(* IEC 61131-3 sources: plcassist-cli/packages/volt-lsp-iec/test-corpus/lenze-mid/Device/Plc Logic/Application/Library Manager/CAA MemBlockMan, 91 files *)

(* ---- RSHANDLING.gvl ---- *)
VAR_GLOBAL
	G_XCHGCLASS : XChgClass;
	G_FLATCLASS : FlatClass;
	G_MSGCLASS : MsgClass;
	G_REFCLASS : MsgClass;
	G_POOLCLASS : PoolClass;
	G_BLKCLASS : BlkClass;
	G_RLSTCLASS : RLstClass;
END_VAR

(* ---- VERSIONCONSTANTS.gvl ---- *)
VAR_GLOBAL
	GC_BYVERSION : BYTE := 1;
	GC_VERSION_1 : BYTE := 0;
END_VAR

(* ---- _BLOCKGETDATA.fun ---- *)
FUNCTION _BLOCKGETDATA : CAA.PVOID
VAR_INPUT
	HBLOCK : CAA.HANDLE;
	PEERROR : POINTER TO ERROR;
END_VAR
END_FUNCTION

(* ---- _BLOCKGETPOOL.fun ---- *)
FUNCTION _BLOCKGETPOOL : CAA.HANDLE
VAR_INPUT
	HBLOCK : CAA.HANDLE;
	PEERROR : POINTER TO ERROR;
END_VAR
END_FUNCTION

(* ---- _FLATCREATEH.fun ---- *)
FUNCTION _FLATCREATEH : CAA.HANDLE
VAR_INPUT
	IDMINKEY : CAA.IDENT;
	IDMAXKEY : CAA.IDENT;
	CTNUMKEYS : CAA.COUNT;
	EENABLE : CB.EVENT;
	EDISABLE : CB.EVENT;
	EUPDATE : CB.EVENT;
	EREAD : CB.EVENT;
	PEERROR : POINTER TO ERROR;
END_VAR
END_FUNCTION

(* ---- _FLATCREATEP.fun ---- *)
FUNCTION _FLATCREATEP : CAA.HANDLE
VAR_INPUT
	IDMINKEY : CAA.IDENT;
	IDMAXKEY : CAA.IDENT;
	CTNUMKEY : CAA.COUNT;
	SZMEMSIZE : CAA.SIZE;
	PMEMORY : CAA.PVOID;
	EENABLE : CB.EVENT;
	EDISABLE : CB.EVENT;
	EUPDATE : CB.EVENT;
	EREAD : CB.EVENT;
	PEERROR : POINTER TO ERROR;
END_VAR
END_FUNCTION

(* ---- _FLATDELETE.fun ---- *)
FUNCTION _FLATDELETE : ERROR
VAR_INPUT
	HFLAT : CAA.HANDLE;
END_VAR
END_FUNCTION

(* ---- _FLATDISABLE.fun ---- *)
FUNCTION _FLATDISABLE : CAA.HANDLE
VAR_INPUT
	HFLAT : CAA.HANDLE;
	IDKEY : CAA.IDENT;
	PEERROR : POINTER TO ERROR;
END_VAR
END_FUNCTION

(* ---- _FLATENABLE.fun ---- *)
FUNCTION _FLATENABLE : ERROR
VAR_INPUT
	HFLAT : CAA.HANDLE;
	IDKEY : CAA.IDENT;
END_VAR
END_FUNCTION

(* ---- _FLATGETSIZE.fun ---- *)
FUNCTION _FLATGETSIZE : CAA.SIZE
VAR_INPUT
	CTNUMKEYS : CAA.COUNT;
END_VAR
END_FUNCTION

(* ---- _FLATREAD.fun ---- *)
FUNCTION _FLATREAD : CAA.HANDLE
VAR_INPUT
	HFLAT : CAA.HANDLE;
	IDKEY : CAA.IDENT;
	PEERROR : POINTER TO ERROR;
END_VAR
END_FUNCTION

(* ---- _FLATTEST.fun ---- *)
FUNCTION _FLATTEST : BOOL
VAR_INPUT
	HFLAT : CAA.HANDLE;
	IDKEY : CAA.IDENT;
	PEERROR : POINTER TO ERROR;
END_VAR
END_FUNCTION

(* ---- _FLATUPDATE.fun ---- *)
FUNCTION _FLATUPDATE : CAA.HANDLE
VAR_INPUT
	HFLAT : CAA.HANDLE;
	IDKEY : CAA.IDENT;
	HMSG : CAA.HANDLE;
	PEERROR : POINTER TO ERROR;
END_VAR
END_FUNCTION

(* ---- _MSGADDREF.fun ---- *)
FUNCTION _MSGADDREF : ERROR
VAR_INPUT
	HMSG : CAA.HANDLE;
END_VAR
END_FUNCTION

(* ---- _MSGCLONE.fun ---- *)
FUNCTION _MSGCLONE : CAA.HANDLE
VAR_INPUT
	HMSG : CAA.HANDLE;
	PEERROR : POINTER TO ERROR;
END_VAR
END_FUNCTION

(* ---- _MSGGETDATA.fun ---- *)
FUNCTION _MSGGETDATA : CAA.PVOID
VAR_INPUT
	HMSG : CAA.HANDLE;
	PEERROR : POINTER TO ERROR;
END_VAR
END_FUNCTION

(* ---- _MSGRECEIVE.fun ---- *)
FUNCTION _MSGRECEIVE : CAA.HANDLE
VAR_INPUT
	HXCHG : CAA.HANDLE;
	PCTMSGLEFT : POINTER TO CAA.COUNT;
	PEERROR : POINTER TO ERROR;
END_VAR
END_FUNCTION

(* ---- _MSGRELEASE.fun ---- *)
FUNCTION _MSGRELEASE : ERROR
VAR_INPUT
	HMSG : CAA.HANDLE;
END_VAR
END_FUNCTION

(* ---- _MSGRELEASEEX.fun ---- *)
FUNCTION _MSGRELEASEEX : ERROR
VAR_INPUT
	HMSG : CAA.HANDLE;
	HXCHG : CAA.HANDLE;
END_VAR
END_FUNCTION

(* ---- _MSGSEND.fun ---- *)
FUNCTION _MSGSEND : ERROR
VAR_INPUT
	HMSG : CAA.HANDLE;
	USIPRIO : USINT;
	HXCHG : CAA.HANDLE;
END_VAR
END_FUNCTION

(* ---- _POOLCREATEH.fun ---- *)
FUNCTION _POOLCREATEH : CAA.HANDLE
VAR_INPUT
	CTNUMBLOCKS : CAA.COUNT;
	SZBLOCKSIZE : CAA.SIZE;
	EEMPTY : CB.EVENT;
	PEERROR : POINTER TO ERROR;
END_VAR
END_FUNCTION

(* ---- _POOLCREATEP.fun ---- *)
FUNCTION _POOLCREATEP : CAA.HANDLE
VAR_INPUT
	SZBLOCKSIZE : CAA.SIZE;
	SZMEMSIZE : CAA.SIZE;
	PMEMORY : CAA.PVOID;
	EEMPTY : CB.EVENT;
	PEERROR : POINTER TO ERROR;
END_VAR
END_FUNCTION

(* ---- _POOLDELETE.fun ---- *)
FUNCTION _POOLDELETE : ERROR
VAR_INPUT
	HPOOL : CAA.HANDLE;
END_VAR
END_FUNCTION

(* ---- _POOLEXTENDH.fun ---- *)
FUNCTION _POOLEXTENDH : ERROR
VAR_INPUT
	HPOOL : CAA.HANDLE;
	CTNUMBLOCKS : CAA.COUNT;
END_VAR
END_FUNCTION

(* ---- _POOLGETBLOCK.fun ---- *)
FUNCTION _POOLGETBLOCK : CAA.HANDLE
VAR_INPUT
	HPOOL : CAA.HANDLE;
	PEERROR : POINTER TO ERROR;
END_VAR
END_FUNCTION

(* ---- _POOLGETBLOCKSIZE.fun ---- *)
FUNCTION _POOLGETBLOCKSIZE : CAA.SIZE
VAR_INPUT
	HPOOL : CAA.HANDLE;
	PEERROR : POINTER TO ERROR;
END_VAR
END_FUNCTION

(* ---- _POOLGETCURCAPACITY.fun ---- *)
FUNCTION _POOLGETCURCAPACITY : CAA.COUNT
VAR_INPUT
	HPOOL : CAA.HANDLE;
	PEERROR : POINTER TO ERROR;
END_VAR
END_FUNCTION

(* ---- _POOLGETNUMBLOCKSLEFT.fun ---- *)
FUNCTION _POOLGETNUMBLOCKSLEFT : CAA.COUNT
VAR_INPUT
	HPOOL : CAA.HANDLE;
	PEERROR : POINTER TO ERROR;
END_VAR
END_FUNCTION

(* ---- _POOLGETSIZE.fun ---- *)
FUNCTION _POOLGETSIZE : CAA.SIZE
VAR_INPUT
	CTNUMBLOCK : CAA.COUNT;
	SZBLOCKSIZE : CAA.SIZE;
END_VAR
END_FUNCTION

(* ---- _POOLPUTBLOCK.fun ---- *)
FUNCTION _POOLPUTBLOCK : ERROR
VAR_INPUT
	HBLOCK : CAA.HANDLE;
END_VAR
END_FUNCTION

(* ---- _RLSTADDPRIO.fun ---- *)
FUNCTION _RLSTADDPRIO : ERROR
VAR_INPUT
	HRLST : CAA.HANDLE;
	USIPRIO : USINT;
END_VAR
END_FUNCTION

(* ---- _RLSTCHECKPRIO.fun ---- *)
FUNCTION _RLSTCHECKPRIO : BOOL
VAR_INPUT
	HRLST : CAA.HANDLE;
	USIPRIO : USINT;
	PEERROR : POINTER TO ERROR;
END_VAR
END_FUNCTION

(* ---- _RLSTCREATEH.fun ---- *)
FUNCTION _RLSTCREATEH : CAA.HANDLE
VAR_INPUT
	PEERROR : POINTER TO ERROR;
END_VAR
END_FUNCTION

(* ---- _RLSTCREATEP.fun ---- *)
FUNCTION _RLSTCREATEP : CAA.HANDLE
VAR_INPUT
	SZMEMORY : CAA.SIZE;
	PMEMORY : CAA.PVOID;
	PEERROR : POINTER TO ERROR;
END_VAR
END_FUNCTION

(* ---- _RLSTDELETE.fun ---- *)
FUNCTION _RLSTDELETE : ERROR
VAR_INPUT
	HRLST : CAA.HANDLE;
END_VAR
END_FUNCTION

(* ---- _RLSTGETHIGHESTPRIO.fun ---- *)
FUNCTION _RLSTGETHIGHESTPRIO : USINT
VAR_INPUT
	HRLST : CAA.HANDLE;
	PEERROR : POINTER TO ERROR;
END_VAR
END_FUNCTION

(* ---- _RLSTGETSIZE.fun ---- *)
FUNCTION _RLSTGETSIZE : CAA.SIZE
VAR_INPUT
	XDUMMY : BOOL;
END_VAR
END_FUNCTION

(* ---- _RLSTREMOVEPRIO.fun ---- *)
FUNCTION _RLSTREMOVEPRIO : ERROR
VAR_INPUT
	HRLST : CAA.HANDLE;
	USIPRIO : USINT;
END_VAR
END_FUNCTION

(* ---- _XCHGCREATEH.fun ---- *)
FUNCTION _XCHGCREATEH : CAA.HANDLE
VAR_INPUT
	CTNUMMSG : CAA.COUNT;
	SZBLOCKSIZE : CAA.SIZE;
	CTNUMPRIOS : CAA.COUNT;
	ESENDMSG : CB.EVENT;
	ERECEIVEMSG : CB.EVENT;
	EXCHGEMPTY : CB.EVENT;
	PEERROR : POINTER TO ERROR;
END_VAR
END_FUNCTION

(* ---- _XCHGCREATEP.fun ---- *)
FUNCTION _XCHGCREATEP : CAA.HANDLE
VAR_INPUT
	SZBLOCKSIZE : CAA.SIZE;
	CTNUMPRIOS : CAA.COUNT;
	SZMEMSIZE : CAA.SIZE;
	PMEMORY : CAA.PVOID;
	ESENDMSG : CB.EVENT;
	ERECEIVEMSG : CB.EVENT;
	EXCHGEMPTY : CB.EVENT;
	PEERROR : POINTER TO ERROR;
END_VAR
END_FUNCTION

(* ---- _XCHGDELETE.fun ---- *)
FUNCTION _XCHGDELETE : ERROR
VAR_INPUT
	HXCHG : CAA.HANDLE;
END_VAR
END_FUNCTION

(* ---- _XCHGEXTENDH.fun ---- *)
FUNCTION _XCHGEXTENDH : ERROR
VAR_INPUT
	HXCHG : CAA.HANDLE;
	CTNUMMSG : CAA.COUNT;
END_VAR
END_FUNCTION

(* ---- _XCHGGETSIZE.fun ---- *)
FUNCTION _XCHGGETSIZE : CAA.SIZE
VAR_INPUT
	CTNUMMSG : CAA.COUNT;
	SZBLOCKSIZE : CAA.SIZE;
	CTNUMPRIOS : CAA.COUNT;
END_VAR
END_FUNCTION

(* ---- _XCHGISEMPTY.fun ---- *)
FUNCTION _XCHGISEMPTY : BOOL
VAR_INPUT
	HXCHG : CAA.HANDLE;
	PEERROR : POINTER TO ERROR;
END_VAR
END_FUNCTION

(* ---- _XCHGMSGLEFT.fun ---- *)
FUNCTION _XCHGMSGLEFT : CAA.COUNT
VAR_INPUT
	HXCHG : CAA.HANDLE;
	PEERROR : POINTER TO ERROR;
END_VAR
END_FUNCTION

(* ---- BLOCKGETDATA.fun ---- *)
FUNCTION BLOCKGETDATA : CAA.PVOID
VAR_INPUT
	HBLOCK : CAA.HANDLE;
	PEERROR : POINTER TO ERROR;
END_VAR
END_FUNCTION

(* ---- FLATCREATEH.fun ---- *)
FUNCTION FLATCREATEH : CAA.HANDLE
VAR_INPUT
	IDMINKEY : CAA.IDENT;
	IDMAXKEY : CAA.IDENT;
	CTNUMKEYS : CAA.COUNT;
	EENABLE : CB.EVENT;
	EDISABLE : CB.EVENT;
	EUPDATE : CB.EVENT;
	EREAD : CB.EVENT;
	PEERROR : POINTER TO ERROR;
END_VAR
END_FUNCTION

(* ---- FLATCREATEP.fun ---- *)
FUNCTION FLATCREATEP : CAA.HANDLE
VAR_INPUT
	IDMINKEY : CAA.IDENT;
	IDMAXKEY : CAA.IDENT;
	CTNUMKEY : CAA.COUNT;
	SZMEMSIZE : CAA.SIZE;
	PMEMORY : CAA.PVOID;
	EENABLE : CB.EVENT;
	EDISABLE : CB.EVENT;
	EUPDATE : CB.EVENT;
	EREAD : CB.EVENT;
	PEERROR : POINTER TO ERROR;
END_VAR
END_FUNCTION

(* ---- FLATDELETE.fun ---- *)
FUNCTION FLATDELETE : ERROR
VAR_INPUT
	HFLAT : CAA.HANDLE;
END_VAR
END_FUNCTION

(* ---- FLATDISABLE.fun ---- *)
FUNCTION FLATDISABLE : CAA.HANDLE
VAR_INPUT
	HFLAT : CAA.HANDLE;
	IDKEY : CAA.IDENT;
	PEERROR : POINTER TO ERROR;
END_VAR
END_FUNCTION

(* ---- FLATENABLE.fun ---- *)
FUNCTION FLATENABLE : ERROR
VAR_INPUT
	HFLAT : CAA.HANDLE;
	IDKEY : CAA.IDENT;
END_VAR
END_FUNCTION

(* ---- FLATGETSIZE.fun ---- *)
FUNCTION FLATGETSIZE : CAA.SIZE
VAR_INPUT
	CTNUMKEYS : CAA.COUNT;
END_VAR
END_FUNCTION

(* ---- FLATREAD.fun ---- *)
FUNCTION FLATREAD : CAA.HANDLE
VAR_INPUT
	HFLAT : CAA.HANDLE;
	IDKEY : CAA.IDENT;
	PEERROR : POINTER TO ERROR;
END_VAR
END_FUNCTION

(* ---- FLATTEST.fun ---- *)
FUNCTION FLATTEST : BOOL
VAR_INPUT
	HFLAT : CAA.HANDLE;
	IDKEY : CAA.IDENT;
	PEERROR : POINTER TO ERROR;
END_VAR
END_FUNCTION

(* ---- FLATUPDATE.fun ---- *)
FUNCTION FLATUPDATE : CAA.HANDLE
VAR_INPUT
	HFLAT : CAA.HANDLE;
	IDKEY : CAA.IDENT;
	HMSG : CAA.HANDLE;
	PEERROR : POINTER TO ERROR;
END_VAR
END_FUNCTION

(* ---- GETSUPPLIERVERSION.fun ---- *)
FUNCTION GETSUPPLIERVERSION : WORD
VAR_INPUT
	XDUMMY : BOOL;
END_VAR
END_FUNCTION

(* ---- MSGADDREF.fun ---- *)
FUNCTION MSGADDREF : ERROR
VAR_INPUT
	HMSG : CAA.HANDLE;
END_VAR
END_FUNCTION

(* ---- MSGCLONE.fun ---- *)
FUNCTION MSGCLONE : CAA.HANDLE
VAR_INPUT
	HMSG : CAA.HANDLE;
	PEERROR : POINTER TO ERROR;
END_VAR
END_FUNCTION

(* ---- MSGGETDATA.fun ---- *)
FUNCTION MSGGETDATA : CAA.PVOID
VAR_INPUT
	HMSG : CAA.HANDLE;
	PEERROR : POINTER TO ERROR;
END_VAR
END_FUNCTION

(* ---- MSGRECEIVE.fun ---- *)
FUNCTION MSGRECEIVE : CAA.HANDLE
VAR_INPUT
	HXCHG : CAA.HANDLE;
	PCTMSGLEFT : POINTER TO CAA.COUNT;
	PEERROR : POINTER TO ERROR;
END_VAR
END_FUNCTION

(* ---- MSGRELEASE.fun ---- *)
FUNCTION MSGRELEASE : ERROR
VAR_INPUT
	HMSG : CAA.HANDLE;
END_VAR
END_FUNCTION

(* ---- MSGRELEASEEX.fun ---- *)
FUNCTION MSGRELEASEEX : ERROR
VAR_INPUT
	HMSG : CAA.HANDLE;
	HXCHG : CAA.HANDLE;
END_VAR
END_FUNCTION

(* ---- MSGSEND.fun ---- *)
FUNCTION MSGSEND : ERROR
VAR_INPUT
	HMSG : CAA.HANDLE;
	USIPRIO : USINT;
	HXCHG : CAA.HANDLE;
END_VAR
END_FUNCTION

(* ---- POOLCREATEH.fun ---- *)
FUNCTION POOLCREATEH : CAA.HANDLE
VAR_INPUT
	CTNUMBLOCKS : CAA.COUNT;
	SZBLOCKSIZE : CAA.SIZE;
	EEMPTY : CB.EVENT;
	PEERROR : POINTER TO ERROR;
END_VAR
END_FUNCTION

(* ---- POOLCREATEP.fun ---- *)
FUNCTION POOLCREATEP : CAA.HANDLE
VAR_INPUT
	SZBLOCKSIZE : CAA.SIZE;
	SZMEMSIZE : CAA.SIZE;
	PMEMORY : CAA.PVOID;
	EEMPTY : CB.EVENT;
	PEERROR : POINTER TO ERROR;
END_VAR
END_FUNCTION

(* ---- POOLDELETE.fun ---- *)
FUNCTION POOLDELETE : ERROR
VAR_INPUT
	HPOOL : CAA.HANDLE;
END_VAR
END_FUNCTION

(* ---- POOLEXTENDH.fun ---- *)
FUNCTION POOLEXTENDH : ERROR
VAR_INPUT
	HPOOL : CAA.HANDLE;
	CTNUMBLOCKS : CAA.COUNT;
END_VAR
END_FUNCTION

(* ---- POOLGETBLOCK.fun ---- *)
FUNCTION POOLGETBLOCK : CAA.HANDLE
VAR_INPUT
	HPOOL : CAA.HANDLE;
	PEERROR : POINTER TO ERROR;
END_VAR
END_FUNCTION

(* ---- POOLGETSIZE.fun ---- *)
FUNCTION POOLGETSIZE : CAA.SIZE
VAR_INPUT
	CTNUMBLOCK : CAA.COUNT;
	SZBLOCKSIZE : CAA.SIZE;
END_VAR
END_FUNCTION

(* ---- POOLPUTBLOCK.fun ---- *)
FUNCTION POOLPUTBLOCK : ERROR
VAR_INPUT
	HBLOCK : CAA.HANDLE;
END_VAR
END_FUNCTION

(* ---- RLSTADDPRIO.fun ---- *)
FUNCTION RLSTADDPRIO : ERROR
VAR_INPUT
	HRLST : CAA.HANDLE;
	USIPRIO : USINT;
END_VAR
END_FUNCTION

(* ---- RLSTCHECKPRIO.fun ---- *)
FUNCTION RLSTCHECKPRIO : BOOL
VAR_INPUT
	HRLST : CAA.HANDLE;
	USIPRIO : USINT;
	PEERROR : POINTER TO ERROR;
END_VAR
END_FUNCTION

(* ---- RLSTCREATEH.fun ---- *)
FUNCTION RLSTCREATEH : CAA.HANDLE
VAR_INPUT
	PEERROR : POINTER TO ERROR;
END_VAR
END_FUNCTION

(* ---- RLSTCREATEP.fun ---- *)
FUNCTION RLSTCREATEP : CAA.HANDLE
VAR_INPUT
	SZMEMORY : CAA.SIZE;
	PMEMORY : CAA.PVOID;
	PEERROR : POINTER TO ERROR;
END_VAR
END_FUNCTION

(* ---- RLSTDELETE.fun ---- *)
FUNCTION RLSTDELETE : ERROR
VAR_INPUT
	HRLST : CAA.HANDLE;
END_VAR
END_FUNCTION

(* ---- RLSTGETHIGHESTPRIO.fun ---- *)
FUNCTION RLSTGETHIGHESTPRIO : USINT
VAR_INPUT
	HRLST : CAA.HANDLE;
	PEERROR : POINTER TO ERROR;
END_VAR
END_FUNCTION

(* ---- RLSTGETSIZE.fun ---- *)
FUNCTION RLSTGETSIZE : CAA.SIZE
VAR_INPUT
	XDUMMY : BOOL;
END_VAR
END_FUNCTION

(* ---- RLSTREMOVEPRIO.fun ---- *)
FUNCTION RLSTREMOVEPRIO : ERROR
VAR_INPUT
	HRLST : CAA.HANDLE;
	USIPRIO : USINT;
END_VAR
END_FUNCTION

(* ---- XCHGCREATEH.fun ---- *)
FUNCTION XCHGCREATEH : CAA.HANDLE
VAR_INPUT
	CTNUMMSG : CAA.COUNT;
	SZBLOCKSIZE : CAA.SIZE;
	CTNUMPRIOS : CAA.COUNT;
	ESENDMSG : CB.EVENT;
	ERECEIVEMSG : CB.EVENT;
	EXCHGEMPTY : CB.EVENT;
	PEERROR : POINTER TO ERROR;
END_VAR
END_FUNCTION

(* ---- XCHGCREATEP.fun ---- *)
FUNCTION XCHGCREATEP : CAA.HANDLE
VAR_INPUT
	SZBLOCKSIZE : CAA.SIZE;
	CTNUMPRIOS : CAA.COUNT;
	SZMEMSIZE : CAA.SIZE;
	PMEMORY : CAA.PVOID;
	ESENDMSG : CB.EVENT;
	ERECEIVEMSG : CB.EVENT;
	EXCHGEMPTY : CB.EVENT;
	PEERROR : POINTER TO ERROR;
END_VAR
END_FUNCTION

(* ---- XCHGDELETE.fun ---- *)
FUNCTION XCHGDELETE : ERROR
VAR_INPUT
	HXCHG : CAA.HANDLE;
END_VAR
END_FUNCTION

(* ---- XCHGEXTENDH.fun ---- *)
FUNCTION XCHGEXTENDH : ERROR
VAR_INPUT
	HXCHG : CAA.HANDLE;
	CTNUMMSG : CAA.COUNT;
END_VAR
END_FUNCTION

(* ---- XCHGGETSIZE.fun ---- *)
FUNCTION XCHGGETSIZE : CAA.SIZE
VAR_INPUT
	CTNUMMSG : CAA.COUNT;
	SZBLOCKSIZE : CAA.SIZE;
	CTNUMPRIOS : CAA.COUNT;
END_VAR
END_FUNCTION

(* ---- XCHGISEMPTY.fun ---- *)
FUNCTION XCHGISEMPTY : BOOL
VAR_INPUT
	HXCHG : CAA.HANDLE;
	PEERROR : POINTER TO ERROR;
END_VAR
END_FUNCTION

(* ---- XCHGMSGLEFT.fun ---- *)
FUNCTION XCHGMSGLEFT : CAA.COUNT
VAR_INPUT
	HXCHG : CAA.HANDLE;
	PEERROR : POINTER TO ERROR;
END_VAR
END_FUNCTION

(* ---- BLKCLASS.fb ---- *)
FUNCTION_BLOCK BLKCLASS EXTENDS RSMClass
END_FUNCTION_BLOCK

METHOD CLOSE : RSM.ERROR
VAR_INPUT
	HHANDLE : CAA.HANDLE;
END_VAR
END_METHOD

(* ---- FLATCLASS.fb ---- *)
FUNCTION_BLOCK FLATCLASS EXTENDS RSMClass
END_FUNCTION_BLOCK

METHOD CLOSE : RSM.ERROR
VAR_INPUT
	HHANDLE : CAA.HANDLE;
END_VAR
END_METHOD

(* ---- MSGCLASS.fb ---- *)
FUNCTION_BLOCK MSGCLASS EXTENDS RSMClass
END_FUNCTION_BLOCK

METHOD CLOSE : RSM.ERROR
VAR_INPUT
	HHANDLE : CAA.HANDLE;
END_VAR
END_METHOD

(* ---- POOLCLASS.fb ---- *)
FUNCTION_BLOCK POOLCLASS EXTENDS RSMClass
END_FUNCTION_BLOCK

METHOD CLOSE : RSM.ERROR
VAR_INPUT
	HHANDLE : CAA.HANDLE;
END_VAR
END_METHOD

(* ---- RLSTCLASS.fb ---- *)
FUNCTION_BLOCK RLSTCLASS EXTENDS RSMClass
END_FUNCTION_BLOCK

METHOD CLOSE : RSM.ERROR
VAR_INPUT
	HHANDLE : CAA.HANDLE;
END_VAR
END_METHOD

(* ---- XCHGCLASS.fb ---- *)
FUNCTION_BLOCK XCHGCLASS EXTENDS RSMClass
END_FUNCTION_BLOCK

METHOD CLOSE : RSM.ERROR
VAR_INPUT
	HHANDLE : CAA.HANDLE;
END_VAR
END_METHOD
